ORGANIZATION_BLOCK "OB_main"
TITLE = "Cyclic interrupt, 100ms"
{ S7_Optimized_Access := 'TRUE' }
VERSION : 0.1

BEGIN
	"Main_DB"();
END_ORGANIZATION_BLOCK
